(* CODESYS project Visu_Prog.export

Project tree, tasks and I/O mapping:
  visualisation Visu_Prog
*)

// /Visu_Prog
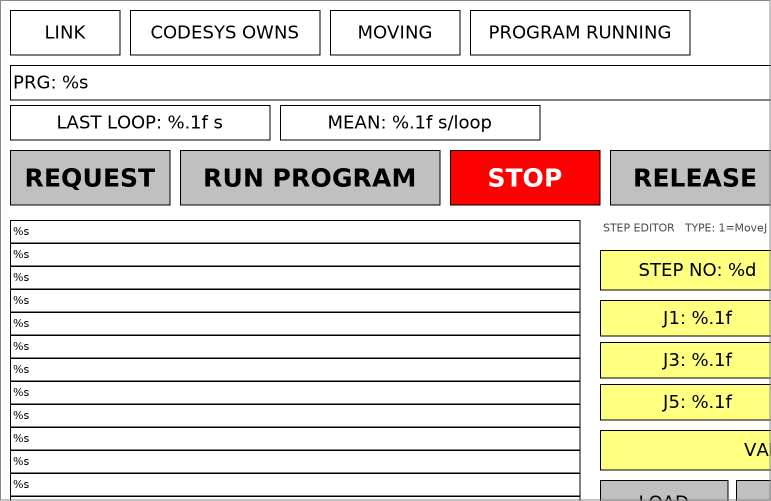
VISUALIZATION Visu_Prog  // 771x501
    Rectangle (10,10 110x45), "LINK", tooltip "Green = Pi and Arduino are talking", colour toggle: P_Arm.xLinkOK
    Rectangle (130,10 190x45), "CODESYS OWNS", tooltip "Green = CODESYS has control of the arm", colour toggle: P_Arm.xOwner
    Rectangle (330,10 130x45), "MOVING", tooltip "Arm is moving", colour toggle: P_Arm.xMoving
    Rectangle (470,10 220x45), "PROGRAM RUNNING", tooltip "Block program is running", colour toggle: P_Arm.xPrgRun
    Rectangle (830,10 170x45), "< ARM PAGE", tooltip "Back to Visu_Arm"
    Rectangle (10,65 990x35), "PRG: %s", tooltip "READY / RUNNING step k/n loop i/N / DONE / STOPPED / ABORTED", text variable: P_Arm.sPrg
    Rectangle (10,105 260x35), "LAST LOOP: %.1f s", tooltip "Time of the last loop", text variable: P_Arm.lrPrgLoopT
    Rectangle (280,105 260x35), "MEAN: %.1f s/loop", tooltip "Mean time per loop", text variable: P_Arm.lrPrgLoopMean
    Rectangle (10,150 160x55), "REQUEST", tooltip "Take control (press before RUN)"
        toggle P_Arm.xBtnRequest
    Rectangle (180,150 260x55), "RUN PROGRAM", tooltip "Run from step 1 to the end"
        toggle P_Arm.xBtnPrgRun
    Rectangle (450,150 150x55), "STOP", tooltip "Stop arm and program now"
        toggle P_Arm.xBtnStop
    Rectangle (610,150 170x55), "RELEASE", tooltip "Give control back to the PC app"
        toggle P_Arm.xBtnRelease
    Rectangle (10,220 570x23), "%s", tooltip "Step 1", text variable: P_Arm.asPrgText[1]
    Rectangle (10,243 570x23), "%s", tooltip "Step 2", text variable: P_Arm.asPrgText[2]
    Rectangle (10,266 570x23), "%s", tooltip "Step 3", text variable: P_Arm.asPrgText[3]
    Rectangle (10,289 570x23), "%s", tooltip "Step 4", text variable: P_Arm.asPrgText[4]
    Rectangle (10,312 570x23), "%s", tooltip "Step 5", text variable: P_Arm.asPrgText[5]
    Rectangle (10,335 570x23), "%s", tooltip "Step 6", text variable: P_Arm.asPrgText[6]
    Rectangle (10,358 570x23), "%s", tooltip "Step 7", text variable: P_Arm.asPrgText[7]
    Rectangle (10,381 570x23), "%s", tooltip "Step 8", text variable: P_Arm.asPrgText[8]
    Rectangle (10,404 570x23), "%s", tooltip "Step 9", text variable: P_Arm.asPrgText[9]
    Rectangle (10,427 570x23), "%s", tooltip "Step 10", text variable: P_Arm.asPrgText[10]
    Rectangle (10,450 570x23), "%s", tooltip "Step 11", text variable: P_Arm.asPrgText[11]
    Rectangle (10,473 570x23), "%s", tooltip "Step 12", text variable: P_Arm.asPrgText[12]
    Rectangle (10,496 570x23), "%s", tooltip "Step 13", text variable: P_Arm.asPrgText[13]
    Rectangle (10,519 570x23), "%s", tooltip "Step 14", text variable: P_Arm.asPrgText[14]
    Rectangle (10,542 570x23), "%s", tooltip "Step 15", text variable: P_Arm.asPrgText[15]
    Rectangle (10,565 570x23), "%s", tooltip "Step 16", text variable: P_Arm.asPrgText[16]
    Rectangle (10,588 570x23), "%s", tooltip "Step 17", text variable: P_Arm.asPrgText[17]
    Rectangle (10,611 570x23), "%s", tooltip "Step 18", text variable: P_Arm.asPrgText[18]
    Rectangle (10,634 570x23), "%s", tooltip "Step 19", text variable: P_Arm.asPrgText[19]
    Rectangle (10,657 570x23), "%s", tooltip "Step 20", text variable: P_Arm.asPrgText[20]
    Label (600,215 400x26), "STEP EDITOR TYPE: 1=MoveJ 2=Speed 3=Wait 4=Loop"
    Rectangle (600,250 195x40), "STEP NO: %d", tooltip "Step to edit 1..20", text variable: P_Arm.iPrgEdit
        OnMouseClick: write the text variable via VisuDialogs.Numpad
    Rectangle (805,250 195x40), "TYPE: %d", tooltip "1=MoveJ 2=Speed 3=Wait 4=Loop", text variable: P_Arm.iEdType
        OnMouseClick: write the text variable via VisuDialogs.Numpad
    Rectangle (600,300 195x36), "J1: %.1f", tooltip "MoveJ angle J1 [deg]", text variable: P_Arm.alrEdJ[0]
        OnMouseClick: write the text variable via VisuDialogs.Numpad
    Rectangle (805,300 195x36), "J2: %.1f", tooltip "MoveJ angle J2 [deg]", text variable: P_Arm.alrEdJ[1]
        OnMouseClick: write the text variable via VisuDialogs.Numpad
    Rectangle (600,342 195x36), "J3: %.1f", tooltip "MoveJ angle J3 [deg]", text variable: P_Arm.alrEdJ[2]
        OnMouseClick: write the text variable via VisuDialogs.Numpad
    Rectangle (805,342 195x36), "J4: %.1f", tooltip "MoveJ angle J4 [deg]", text variable: P_Arm.alrEdJ[3]
        OnMouseClick: write the text variable via VisuDialogs.Numpad
    Rectangle (600,384 195x36), "J5: %.1f", tooltip "MoveJ angle J5 [deg]", text variable: P_Arm.alrEdJ[4]
        OnMouseClick: write the text variable via VisuDialogs.Numpad
    Rectangle (805,384 195x36), "J6: %.1f", tooltip "MoveJ angle J6 [deg]", text variable: P_Arm.alrEdJ[5]
        OnMouseClick: write the text variable via VisuDialogs.Numpad
    Rectangle (600,430 400x40), "VALUE: %.1f", tooltip "Speed [%] / Wait [s] / Loop [count]", text variable: P_Arm.lrEdVal
        OnMouseClick: write the text variable via VisuDialogs.Numpad
    Rectangle (600,480 128x45), "LOAD", tooltip "Load step STEP NO into the editor"
        toggle P_Arm.xBtnPrgLoad
    Rectangle (736,480 128x45), "SAVE", tooltip "Save editor over step STEP NO"
        toggle P_Arm.xBtnPrgSave
    Rectangle (872,480 128x45), "INSERT", tooltip "Insert editor as new step at STEP NO"
        toggle P_Arm.xBtnPrgIns
    Rectangle (600,535 128x45), "DELETE", tooltip "Delete step STEP NO"
        toggle P_Arm.xBtnPrgDel
    Rectangle (736,535 264x45), "TEACH (ACTUAL > J)", tooltip "Copy actual angles into J1..J6"
        toggle P_Arm.xBtnPrgTeach
    Rectangle (600,590 400x40), "DEFAULT PEN PROGRAM", tooltip "Reload the 12-step pen program"
        toggle P_Arm.xBtnPrgDefault
END_VISUALIZATION
